Staubli VAL3: do_endSwitch.pgx

public program do_endSwitch()
begin
  rs:bInSwitch=false
end
